FUNCTION_BLOCK StructScopeTest (* Simple FB validating structured member lookup *)
  (* Standard: 61499-1; Description: Copyright (c) 2026 Martin Erich Jobst This program and the accompanying materials are made available under the terms of the Eclipse Public License 2.0 which is available at https://www.eclipse.org/legal/epl-2.0/ SPDX-License-Identifier: EPL-2.0 *)
  (* Version 1.0, 2026-11-18, Martin Jobst *)
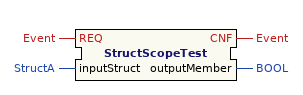
  EVENT_INPUT
    REQ; (* Normal Execution Request *)
  END_EVENT
  EVENT_OUTPUT
    CNF; (* Execution Confirmation *)
  END_EVENT
  VAR_INPUT
    inputStruct : StructA;
  END_VAR
  VAR_OUTPUT
    outputMember : BOOL;
  END_VAR
  EC_STATES
    REQ : REQ -> CNF;
  END_STATES
  ALGORITHM REQ IN ST:
VAR_TEMP
	initializedStruct : StructScopeType := (visibleMember := TRUE, unavailableInitializerMember := FALSE);
END_VAR
initializedStruct.visibleMember := TRUE;
initializedStruct.unavailableReceiverMember := FALSE;
outputMember := initializedStruct.visibleMember;
outputMember := inputStruct.nestedStruct.visibleMember;
  END_ALGORITHM
END_FUNCTION_BLOCK
